TYPE stLightState :
STRUCT
	PowerOn : BOOL;
	Color : stLightColor;
	Temperature : eLightTemperature;
	Brightness : USINT;		// 20 - 100%
END_STRUCT
END_TYPE

(* stored: Version 1.1.0.1
   DUT stLightState: Id {90c9e709-c995-434d-b1ec-c79b08482bcc} *)
